(* CODESYS project SingleElevator.project

Project tree, tasks and I/O mapping:
  Device : CODESYS Control Win V3, 3S - Smart Software Solutions GmbH, version 3.5.18.0
    application Application
      libraries: Standard, 3.5.18.0 (System)
      task MainTask (cyclic, interval t#20ms, priority 1) calls GAs_Collector, Simulation, Policy
      task VISU_TASK (cyclic, interval 100 ms, priority 31) calls VisuElems.Visu_Prg
      global variables GVL
      visualisation Visualization
      program Simulation [ST]
      function block Cabin_GA [SFC]: Init_active, Ready_active, Busy_active, CabinUP_active, CabinUP_exit, CabinDown_exit, CabinDown_active, DoneHoming_active, DoneHoming_exit, HomingUp_active, HomingUp_exit, Step0_active, Step0_exit, ConteggioRampe_active, ConteggioDeck_active, Rallenta_active, Rallenta_exit, Fault_active, DoneCabin_active, FaultDeck_active, FaultDoneD_active, FaultDoneD_exit, FaultRamp_active, FaultDoneR_active, FaultDoneR_exit, FaultLimit_active, FaultLimit_exit, FaultDoneL_active, FaultDoneL_exit
      function block Doors_GA [SFC]: Init_active, Ready_active, Ready_exit, DoorOpening_active, DoorOpening_exit, SetDoneO_active, SetDoneO_exit, DoorClosing_active, DoorClosing_exit, SetDoneC_active, SetDoneC_exit
      function block HMI_GA [SFC]: Init_active, Ready_active, Ready_exit, LED_active, Chiamate_active, Destinazioni_active
      program Policy [SFC]: ChiusuraHoming_active, ChiusuraHoming_exit, Homing_active, Homing_exit, AperturaHoming_active, AperturaHoming_exit, Wait_Call_active, CalcoloDest_active, StopHMI_active, Chiudi_exit, Chiudi_active, Rallenta_active, AperturaEmergenza_active, Sali_active, Scendi_active, Sali_exit, Scendi_exit, Apri_exit, Apri_active
      program GAs_Collector [FBD]
  text list GlobalTextList
*)

// Device/Application/GVL

//{attribute 'qualified_only'}
VAR_GLOBAL
(* Elevator managing variables*)
	Open: BOOL;				(* Sensor: the door is fully open*)
	Closed: BOOL;			(* Sensor: the door is fully closed*)
	LimitDown: BOOL;		(* Sensor: lower limit sensor, if TRUE the lift has reached the lower limit*)
	LimitUp: BOOL;			(* Sensor: upper limit sensor, if TRUE the lift has reached the upper limit*)
	DeckSensor: BOOL;		(* Sensor: if TRUE the cab is in proximity of a deck*)
	RampSensor: BOOL;		(* Sensor: if TRUE the cab is in proximity of a ramp*)
	Presence :BOOL; 		(* Sensor: if TRUE something blocks the door photocell*)
	Emergency: BOOL;		(* Input: if TRUE the emergency button has been pressed*)

	Closing: BOOL;			(* Actuator: if TRUE the door starts closing*)
	Opening: BOOL;			(* Actuator: the door starts opening*)
	Motor_on: BOOL;			(* Actuator: if TRUE the lift pulley motor start moving*)
	Up: BOOL;				(* Actuator parameter: if TRUE the lift moves upward, downward otherwise*)
	Vel: BOOL;				(* Actuator parameter: motor speed, if TRUE high speed, low speed otherwise*)


	Current: INT;  			(* Visualization: variable used to storage the current deck*)
    Destination: INT;		(* Visualization: variable used to storage the the destination deck*)
	EmergencyVis: BOOL; 	(* Visualization: if TRUE the emergency light is turned on*)

	InitialDeck: INT := 1;	(* Only for simulation: variable used to define the initial deck*)
	InitCycle: BOOL := FALSE;(* Only for simulation: used to execute the instruction at the first cycle*)
	Height: INT;			(* Only for simulation: elevator height*)
	DeckRest: INT;        	(* Only for simulation: division rest for generating deck sensor*)
	Memory: INT;
	RampRest: INT;			(* Only for simulation: division rest for generating the ramp position*)
	MemoryR: INT;
	Door: INT;				(* Only for simulation: to visualize the closing of the door*)
	Displacement: INT;		(* Only for simulation: lift displacement, dependent on the motor speed*)

 (*Inputs: internal panel variables*)
	PG: BOOL;
	P1: BOOL;
	P2: BOOL;
	P3: BOOL;
	P4: BOOL;
	P5: BOOL;
	P6: BOOL;
	P7: BOOL;

(*Visualization: internal panel variables used to turn on the LED*)
	PGVis: BOOL;
	P1Vis: BOOL;
	P2Vis: BOOL;
	P3Vis: BOOL;
	P4Vis: BOOL;
	P5Vis: BOOL;
	P6Vis: BOOL;
	P7Vis: BOOL;

(*Inputs: external panel variables*)
	UpDeckG: BOOL;
	UpDeck1: BOOL;
	UpDeck2: BOOL;
	UpDeck3: BOOL;
	UpDeck4: BOOL;
	UpDeck5: BOOL;
	UpDeck6: BOOL;
	DownDeck7: BOOL;
	DownDeck6: BOOL;
	DownDeck5: BOOL;
	DownDeck4: BOOL;
	DownDeck3: BOOL;
	DownDeck2: BOOL;
	DownDeck1: BOOL;

(*Visualization: external panel variables used to turn on the LED*)
	UpDeckGVis: BOOL;
	UpDeck1Vis: BOOL;
	UpDeck2Vis: BOOL;
	UpDeck3Vis: BOOL;
	UpDeck4Vis: BOOL;
	UpDeck5Vis: BOOL;
	UpDeck6Vis: BOOL;
	DownDeck7Vis: BOOL;
	DownDeck6Vis: BOOL;
	DownDeck5Vis: BOOL;
	DownDeck4Vis: BOOL;
	DownDeck3Vis: BOOL;
	DownDeck2Vis: BOOL;
	DownDeck1Vis: BOOL;

(*Only for simulation: variables used to simulate the fault on deck sensor*)
	SensorG: BOOL;				(* if TRUE the magnetic information for deck G is lost and the deck sensor cannot become TRUE*)
	Sensor1: BOOL;				(* if TRUE the magnetic information for deck 1 is lost and the deck sensor cannot become TRUE*)
	Sensor2: BOOL;
	Sensor3: BOOL;
	Sensor4: BOOL;
	Sensor5: BOOL;
	Sensor6: BOOL;
	Sensor7: BOOL;
	FaultSensorAlarm: BOOL; 	(* Visulaization: if TRUE alerts the user of a deck sensor fault*)

(*Only for simulation: variables used to simulate the fault on ramp sensor*)
	RampGUp: BOOL;
	Ramp1Down: BOOL;
	Ramp1Up:BOOL;
	Ramp2Down: BOOL;
	Ramp2Up:BOOL;
	Ramp3Down: BOOL;
	Ramp3Up:BOOL;
	Ramp4Down: BOOL;
	Ramp4Up:BOOL;
	Ramp5Down: BOOL;
	Ramp5Up:BOOL;
	Ramp6Down: BOOL;
	Ramp6Up:BOOL;
	Ramp7Down: BOOL;
	FaultRampAlarm: BOOL; 		(* Visulaization: if TRUE alerts the user of a ramp sensor fault*)
	SensorGOK: BOOL;
	Sensor1OK: BOOL;
	Sensor2OK: BOOL;
	Sensor6OK: BOOL;
	Sensor3OK: BOOL;
	Sensor4OK: BOOL;
	Sensor5OK: BOOL;
	Sensor7OK: BOOL;
	RampGUpOK: BOOL;
	Ramp1DownOK: BOOL;
	Ramp1UpOK: BOOL;
	Ramp2DownOK: BOOL;
	Ramp2UpOK: BOOL;
	Ramp3DownOK: BOOL;
	Ramp3UpOK: BOOL;
	Ramp4DownOK: BOOL;
	Ramp4UpOK: BOOL;
	Ramp5DownOK: BOOL;
	Ramp5UpOK: BOOL;
	Ramp6DownOK: BOOL;
	Ramp6UpOK: BOOL;
	Ramp7DownOK: BOOL;
	Ramp7UpOK: BOOL;
	
	
	Cabin_GA_0: Cabin_GA;
	Doors_GA_0: Doors_GA;
	HMI_GA_0: HMI_GA;
END_VAR

// Device/Application/GAs_Collector
PROGRAM GAs_Collector
VAR
END_VAR

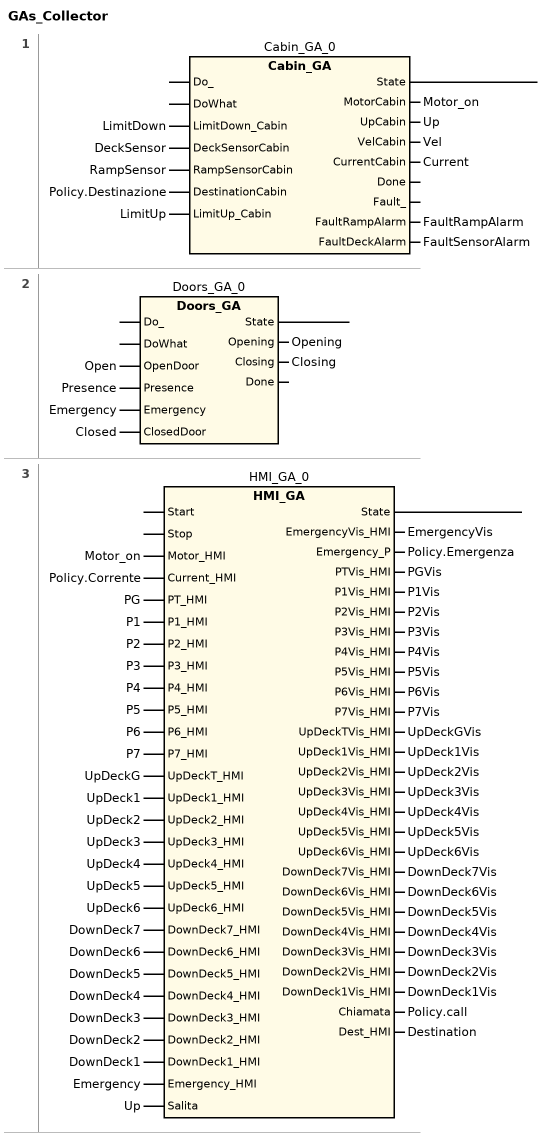
// NETWORK 1
Cabin_GA_0(
    LimitDown_Cabin := LimitDown,
    DeckSensorCabin := DeckSensor,
    RampSensorCabin := RampSensor,
    DestinationCabin := Policy.Destinazione,
    LimitUp_Cabin := LimitUp,
    MotorCabin => Motor_on,
    UpCabin => Up,
    VelCabin => Vel,
    CurrentCabin => Current,
    FaultRampAlarm => FaultRampAlarm,
    FaultDeckAlarm => FaultSensorAlarm); // Cabin_GA

// NETWORK 2
Doors_GA_0(
    OpenDoor := Open,
    Presence := Presence,
    Emergency := Emergency,
    ClosedDoor := Closed,
    Opening => Opening,
    Closing => Closing); // Doors_GA

// NETWORK 3
HMI_GA_0(
    Motor_HMI := Motor_on,
    Current_HMI := Policy.Corrente,
    PT_HMI := PG,
    P1_HMI := P1,
    P2_HMI := P2,
    P3_HMI := P3,
    P4_HMI := P4,
    P5_HMI := P5,
    P6_HMI := P6,
    P7_HMI := P7,
    UpDeckT_HMI := UpDeckG,
    UpDeck1_HMI := UpDeck1,
    UpDeck2_HMI := UpDeck2,
    UpDeck3_HMI := UpDeck3,
    UpDeck4_HMI := UpDeck4,
    UpDeck5_HMI := UpDeck5,
    UpDeck6_HMI := UpDeck6,
    DownDeck7_HMI := DownDeck7,
    DownDeck6_HMI := DownDeck6,
    DownDeck5_HMI := DownDeck5,
    DownDeck4_HMI := DownDeck4,
    DownDeck3_HMI := DownDeck3,
    DownDeck2_HMI := DownDeck2,
    DownDeck1_HMI := DownDeck1,
    Emergency_HMI := Emergency,
    Salita := Up,
    EmergencyVis_HMI => EmergencyVis,
    Emergency_P => Policy.Emergenza,
    PTVis_HMI => PGVis,
    P1Vis_HMI => P1Vis,
    P2Vis_HMI => P2Vis,
    P3Vis_HMI => P3Vis,
    P4Vis_HMI => P4Vis,
    P5Vis_HMI => P5Vis,
    P6Vis_HMI => P6Vis,
    P7Vis_HMI => P7Vis,
    UpDeckTVis_HMI => UpDeckGVis,
    UpDeck1Vis_HMI => UpDeck1Vis,
    UpDeck2Vis_HMI => UpDeck2Vis,
    UpDeck3Vis_HMI => UpDeck3Vis,
    UpDeck4Vis_HMI => UpDeck4Vis,
    UpDeck5Vis_HMI => UpDeck5Vis,
    UpDeck6Vis_HMI => UpDeck6Vis,
    DownDeck7Vis_HMI => DownDeck7Vis,
    DownDeck6Vis_HMI => DownDeck6Vis,
    DownDeck5Vis_HMI => DownDeck5Vis,
    DownDeck4Vis_HMI => DownDeck4Vis,
    DownDeck3Vis_HMI => DownDeck3Vis,
    DownDeck2Vis_HMI => DownDeck2Vis,
    DownDeck1Vis_HMI => DownDeck1Vis,
    Chiamata => Policy.call,
    Dest_HMI => Destination); // HMI_GA

END_PROGRAM

// Device/Application/Cabin_GA
FUNCTION_BLOCK Cabin_GA
VAR_INPUT
	Do_: BOOL;
	DoWhat: STRING;
	LimitDown_Cabin: BOOL;
	DeckSensorCabin: BOOL;
	RampSensorCabin: BOOL;
	DestinationCabin: INT;
	LimitUp_Cabin: BOOL;
END_VAR
VAR_OUTPUT
	State: STRING;
	MotorCabin: BOOL;
	UpCabin: BOOL;
	VelCabin: BOOL;
	CurrentCabin: INT;
	Done: BOOL;
	Fault_: BOOL;
	FaultRampAlarm: BOOL;
	FaultDeckAlarm: BOOL;
END_VAR
VAR
	N_rampe: INT;
	Dest: INT;
	Start: INT;
	i: INT; (*Rampe*)
	j: INT; (*Deck*)
	//k: INT; (*Rampe Aggiuntivo*)
	D_: BOOL;
	R_: BOOL;
	LUC: BOOL;
	LDC: BOOL;
END_VAR

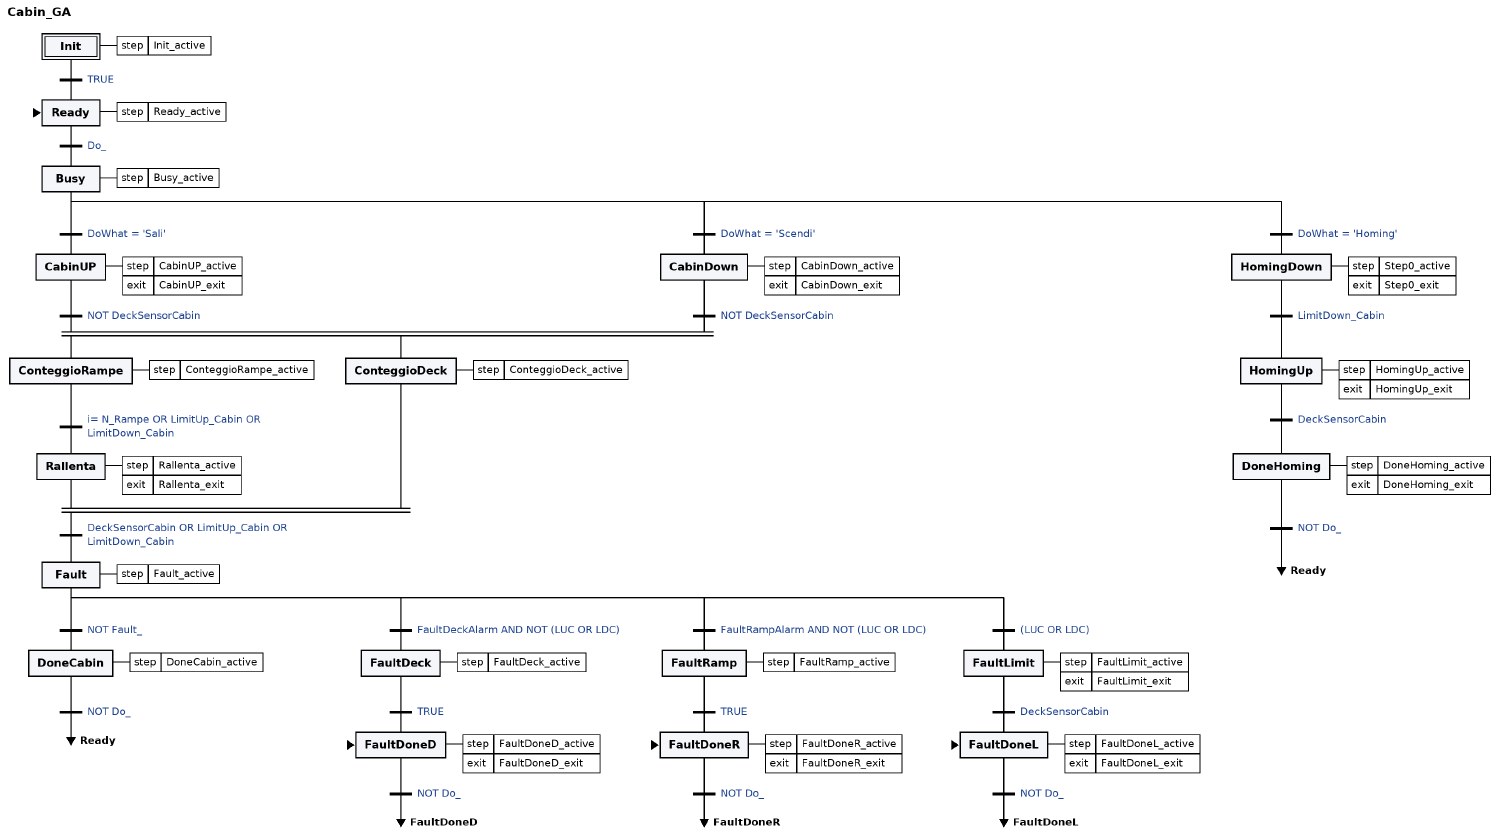
INITIAL_STEP Init:
    Init_active(N);  // step action
END_STEP
TRANSITION FROM Init TO Ready
    := TRUE;
END_TRANSITION
STEP Ready:
    Ready_active(N);  // step action
END_STEP
TRANSITION FROM Ready TO Busy
    := Do_;
END_TRANSITION
STEP Busy:
    Busy_active(N);  // step action
END_STEP
TRANSITION FROM Busy TO CabinUP
    := DoWhat = 'Sali';
END_TRANSITION
STEP CabinUP:
    CabinUP_active(N);  // step action
    CabinUP_exit(P0);  // exit action
END_STEP
TRANSITION FROM CabinUP TO (ConteggioRampe, ConteggioDeck)
    := NOT DeckSensorCabin;
END_TRANSITION
TRANSITION FROM Busy TO CabinDown
    := DoWhat = 'Scendi';
END_TRANSITION
STEP CabinDown:
    CabinDown_active(N);  // step action
    CabinDown_exit(P0);  // exit action
END_STEP
TRANSITION FROM CabinDown TO (ConteggioRampe, ConteggioDeck)
    := NOT DeckSensorCabin;
END_TRANSITION
TRANSITION FROM Busy TO HomingDown
    := DoWhat = 'Homing';
END_TRANSITION
STEP HomingDown:
    Step0_active(N);  // step action
    Step0_exit(P0);  // exit action
END_STEP
TRANSITION FROM HomingDown TO HomingUp
    := LimitDown_Cabin;
END_TRANSITION
STEP HomingUp:
    HomingUp_active(N);  // step action
    HomingUp_exit(P0);  // exit action
END_STEP
TRANSITION FROM HomingUp TO DoneHoming
    := DeckSensorCabin;
END_TRANSITION
STEP DoneHoming:
    DoneHoming_active(N);  // step action
    DoneHoming_exit(P0);  // exit action
END_STEP
TRANSITION FROM DoneHoming TO Ready
    := NOT Do_;
END_TRANSITION
STEP ConteggioRampe:
    ConteggioRampe_active(N);  // step action
END_STEP
TRANSITION FROM ConteggioRampe TO Rallenta
    := i= N_Rampe OR LimitUp_Cabin OR LimitDown_Cabin;
END_TRANSITION
STEP Rallenta:
    Rallenta_active(N);  // step action
    Rallenta_exit(P0);  // exit action
END_STEP
STEP ConteggioDeck:
    ConteggioDeck_active(N);  // step action
END_STEP
TRANSITION FROM (Rallenta, ConteggioDeck) TO Fault
    := DeckSensorCabin OR LimitUp_Cabin OR LimitDown_Cabin;
END_TRANSITION
STEP Fault:
    Fault_active(N);  // step action
END_STEP
TRANSITION FROM Fault TO DoneCabin
    := NOT Fault_;
END_TRANSITION
STEP DoneCabin:
    DoneCabin_active(N);  // step action
END_STEP
TRANSITION FROM DoneCabin TO Ready
    := NOT Do_;
END_TRANSITION
TRANSITION FROM Fault TO FaultDeck
    := FaultDeckAlarm AND NOT (LUC OR LDC);
END_TRANSITION
STEP FaultDeck:
    FaultDeck_active(N);  // step action
END_STEP
TRANSITION FROM FaultDeck TO FaultDoneD
    := TRUE;
END_TRANSITION
STEP FaultDoneD:
    FaultDoneD_active(N);  // step action
    FaultDoneD_exit(P0);  // exit action
END_STEP
TRANSITION FROM FaultDoneD TO FaultDoneD
    := NOT Do_;
END_TRANSITION
TRANSITION FROM Fault TO FaultRamp
    := FaultRampAlarm AND NOT (LUC OR LDC);
END_TRANSITION
STEP FaultRamp:
    FaultRamp_active(N);  // step action
END_STEP
TRANSITION FROM FaultRamp TO FaultDoneR
    := TRUE;
END_TRANSITION
STEP FaultDoneR:
    FaultDoneR_active(N);  // step action
    FaultDoneR_exit(P0);  // exit action
END_STEP
TRANSITION FROM FaultDoneR TO FaultDoneR
    := NOT Do_;
END_TRANSITION
TRANSITION FROM Fault TO FaultLimit
    := (LUC OR LDC);
END_TRANSITION
STEP FaultLimit:
    FaultLimit_active(N);  // step action
    FaultLimit_exit(P0);  // exit action
END_STEP
TRANSITION FROM FaultLimit TO FaultDoneL
    := DeckSensorCabin;
END_TRANSITION
STEP FaultDoneL:
    FaultDoneL_active(N);  // step action
    FaultDoneL_exit(P0);  // exit action
END_STEP
TRANSITION FROM FaultDoneL TO FaultDoneL
    := NOT Do_;
END_TRANSITION

ACTION Init_active:
State := 'Init';
END_ACTION

ACTION Ready_active:
State := 'Ready';
END_ACTION

ACTION Busy_active:
State := 'Busy';
END_ACTION

ACTION CabinUP_active:
MotorCabin := TRUE;
UpCabin := TRUE;
VelCabin :=FALSE;


N_rampe := (ABS(DestinationCabin - CurrentCabin)*2); (*Sensori di rampa attraversati*)
Dest := DestinationCabin;
Start:= CurrentCabin;
i:=0;
j:=0;
END_ACTION

ACTION CabinUP_exit:
VelCabin := TRUE;
END_ACTION

ACTION CabinDown_exit:
VelCabin := TRUE;
END_ACTION

ACTION CabinDown_active:
MotorCabin := TRUE;
UpCabin := FALSE;
VelCabin := FALSE;


N_rampe := (ABS(DestinationCabin - CurrentCabin)*2); (*Sensori di rampa attraversati*)
Dest := DestinationCabin;
Start:= CurrentCabin;
i:=0;
j:=0;
END_ACTION

ACTION DoneHoming_active:
Done :=TRUE;
END_ACTION

ACTION DoneHoming_exit:
Done := FALSE;
END_ACTION

ACTION HomingUp_active:
MotorCabin := TRUE;
UpCabin := TRUE;
VelCabin := FALSE;
END_ACTION

ACTION HomingUp_exit:
MotorCabin := FALSE;
CurrentCabin := 0;
END_ACTION

ACTION Step0_active:
MotorCabin := TRUE;
UpCabin := FALSE;
VelCabin := FALSE;
END_ACTION

ACTION Step0_exit:
MotorCabin := FALSE;
END_ACTION

ACTION ConteggioRampe_active:
IF RampSensorCabin = TRUE THEN
	IF R_ THEN
		i:=i+1;
		R_:=FALSE;
	END_IF
ELSE
	R_:=TRUE;
END_IF


IF Dest <> DestinationCabin THEN
	N_rampe := (ABS(DestinationCabin - Start)*2);
	Dest:=DestinationCabin;
END_IF
END_ACTION

ACTION ConteggioDeck_active:
IF DeckSensorCabin = TRUE THEN
	IF D_ THEN
		j:=j+1;
		D_:=FALSE;
		IF DoWhat = 'Sali' THEN
			CurrentCabin := CurrentCabin+1;
		ELSE
			CurrentCabin := CurrentCabin-1;
		END_IF
	END_IF
ELSE
	D_:=TRUE;
END_IF
END_ACTION

ACTION Rallenta_active:
VelCabin := FALSE;

IF RampSensor=TRUE THEN
	IF R_ THEN
		i:=i+1;
		R_:=FALSE;
	END_IF
ELSE
	R_:=TRUE;
END_IF
END_ACTION

ACTION Rallenta_exit:
MotorCabin := FALSE;
UpCabin := FALSE;
END_ACTION

ACTION Fault_active:
//Fault Deck/Fault Ramp
IF i<(2*j) AND NOT LUC AND NOT LDC THEN
	FaultRampAlarm :=TRUE;
	Fault_:=TRUE;
ELSIF i>(2*j) THEN
	FaultDeckAlarm :=TRUE;
	Fault_:=TRUE;
END_IF

//Fault Limit Up/Limit Down
IF LimitUp_Cabin THEN
	MotorCabin := TRUE;
	UpCabin:=FALSE;
	VelCabin := FALSE;
	LUC :=TRUE;
END_IF

IF LimitDown_Cabin THEN
	MotorCabin := TRUE;
	UpCabin:=TRUE;
	VelCabin := FALSE;
	LDC :=TRUE;
END_IF

IF LUC OR LDC THEN
	Fault_:=TRUE;
END_IF

//No Fault
IF i=2*j THEN
	Fault_:=FALSE;
END_IF
END_ACTION

ACTION DoneCabin_active:
Done := TRUE;
END_ACTION

ACTION FaultDeck_active:
IF DoWhat = 'Sali' THEN
	CurrentCabin := DestinationCabin+1;
ELSIF DoWhat = 'Scendi' THEN
	CurrentCabin := DestinationCabin-1;
END_IF

State := 'Fault_Deck';
DoWhat := 'Stop';
END_ACTION

ACTION FaultDoneD_active:
Done := TRUE;
END_ACTION

ACTION FaultDoneD_exit:
Done := FALSE;
END_ACTION

ACTION FaultRamp_active:
IF DoWhat = 'Sali' THEN
	CurrentCabin := DestinationCabin+1;
ELSIF DoWhat = 'Scendi' THEN
	CurrentCabin := DestinationCabin-1;
END_IF

State := 'Fault_Ramp';
DoWhat := 'Stop';
END_ACTION

ACTION FaultDoneR_active:
Done := TRUE;
END_ACTION

ACTION FaultDoneR_exit:
Done := FALSE;
END_ACTION

ACTION FaultLimit_active:
IF LUC THEN
	State := 'Fault_Deck';
END_IF

IF LDC THEN
	State:= 'Fault_Deck';
END_IF
END_ACTION

ACTION FaultLimit_exit:
MotorCabin := FALSE;
END_ACTION

ACTION FaultDoneL_active:
Done := TRUE;
END_ACTION

ACTION FaultDoneL_exit:
Done := false;
END_ACTION

END_FUNCTION_BLOCK

// Device/Application/Policy
PROGRAM Policy
VAR
	sync: BOOL;
	OpOk: BOOL;
	
	Destinazione: INT;
	Corrente: INT;
END_VAR

VAR_INPUT
	call: BOOL; 					//Presenza chiamate (origine: HMI)
	Emergenza: BOOL;				//Variabile di appoggio per Emergency (origine: HMI)
END_VAR

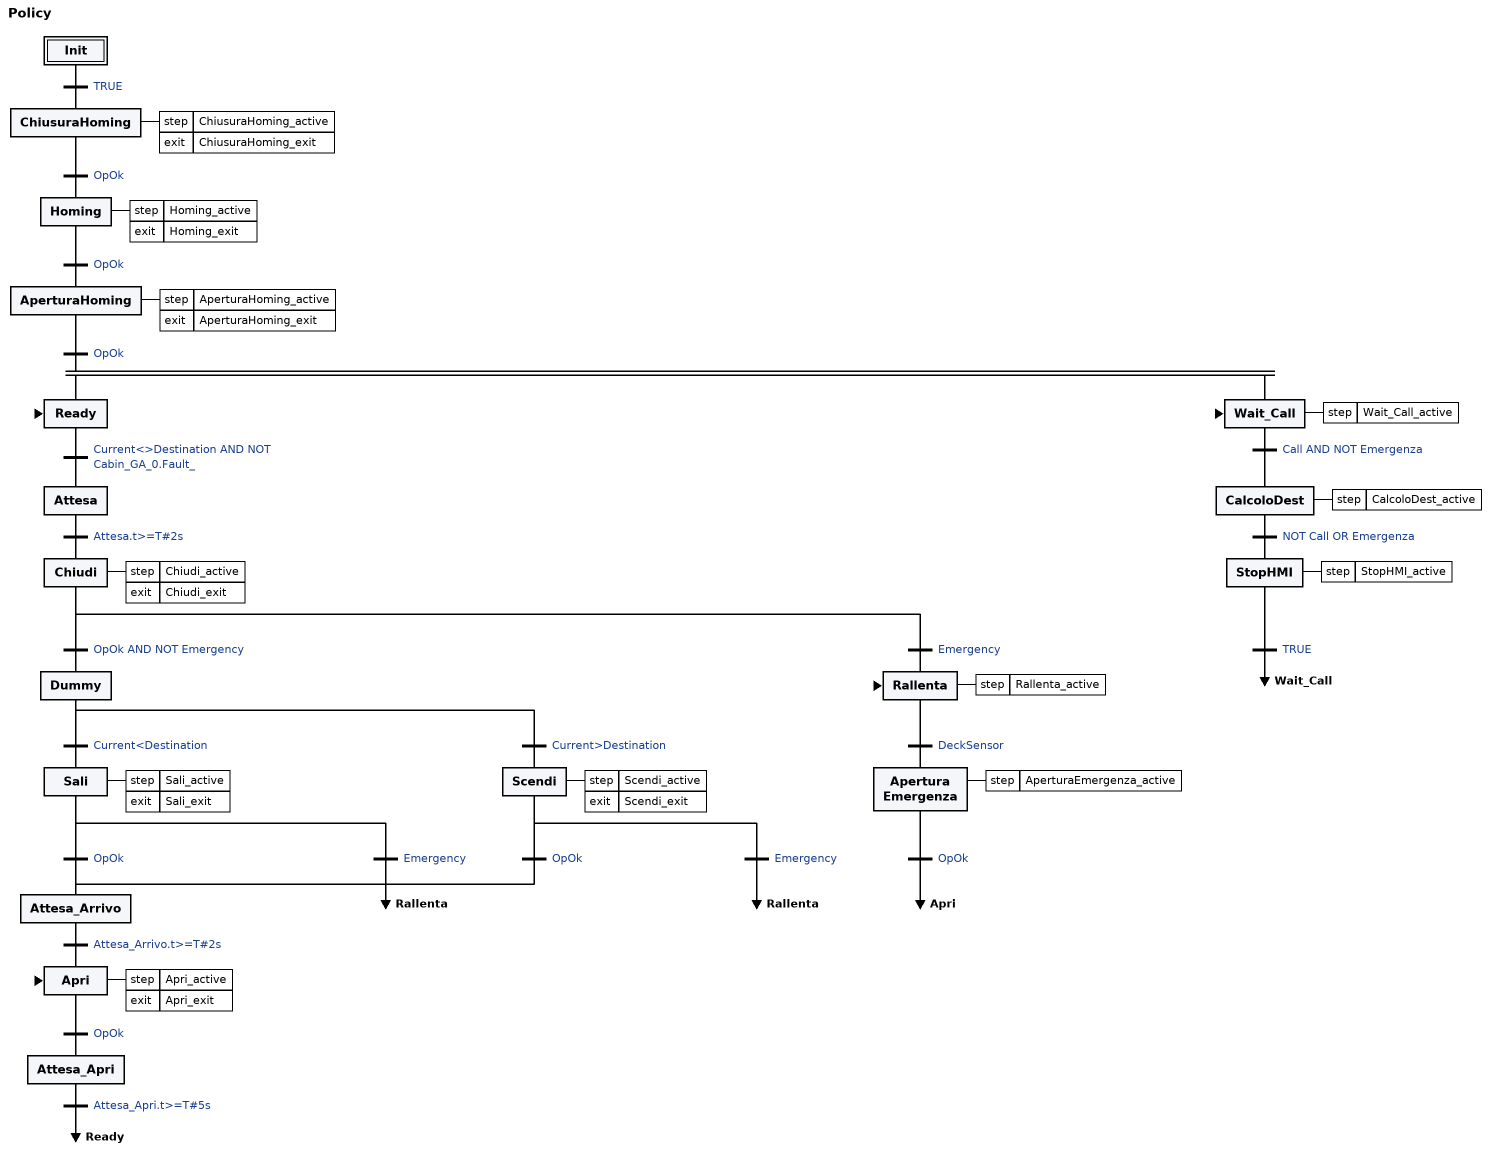
INITIAL_STEP Init:
END_STEP
TRANSITION FROM Init TO ChiusuraHoming
    := TRUE;
END_TRANSITION
STEP ChiusuraHoming:
    ChiusuraHoming_active(N);  // step action
    ChiusuraHoming_exit(P0);  // exit action
END_STEP
TRANSITION FROM ChiusuraHoming TO Homing
    := OpOk;
END_TRANSITION
STEP Homing:
    Homing_active(N);  // step action
    Homing_exit(P0);  // exit action
END_STEP
TRANSITION FROM Homing TO AperturaHoming
    := OpOk;
END_TRANSITION
STEP AperturaHoming:
    AperturaHoming_active(N);  // step action
    AperturaHoming_exit(P0);  // exit action
END_STEP
TRANSITION FROM AperturaHoming TO (Ready, Wait_Call)
    := OpOk;
END_TRANSITION
STEP Ready:
END_STEP
TRANSITION FROM Ready TO Attesa
    := Current<>Destination AND NOT Cabin_GA_0.Fault_;
END_TRANSITION
STEP Attesa:
END_STEP
TRANSITION FROM Attesa TO Chiudi
    := Attesa.t>=T#2s;
END_TRANSITION
STEP Chiudi:
    Chiudi_active(N);  // step action
    Chiudi_exit(P0);  // exit action
END_STEP
TRANSITION FROM Chiudi TO Dummy
    := OpOk AND NOT Emergency;
END_TRANSITION
STEP Dummy:
END_STEP
TRANSITION FROM Dummy TO Sali
    := Current<Destination;
END_TRANSITION
STEP Sali:
    Sali_active(N);  // step action
    Sali_exit(P0);  // exit action
END_STEP
TRANSITION FROM Sali TO Attesa_Arrivo
    := OpOk;
END_TRANSITION
TRANSITION FROM Sali TO Rallenta
    := Emergency;
END_TRANSITION
TRANSITION FROM Dummy TO Scendi
    := Current>Destination;
END_TRANSITION
STEP Scendi:
    Scendi_active(N);  // step action
    Scendi_exit(P0);  // exit action
END_STEP
TRANSITION FROM Scendi TO Attesa_Arrivo
    := OpOk;
END_TRANSITION
TRANSITION FROM Scendi TO Rallenta
    := Emergency;
END_TRANSITION
STEP Attesa_Arrivo:
END_STEP
TRANSITION FROM Attesa_Arrivo TO Apri
    := Attesa_Arrivo.t>=T#2s;
END_TRANSITION
STEP Apri:
    Apri_active(N);  // step action
    Apri_exit(P0);  // exit action
END_STEP
TRANSITION FROM Apri TO Attesa_Apri
    := OpOk;
END_TRANSITION
STEP Attesa_Apri:
END_STEP
TRANSITION FROM Attesa_Apri TO Ready
    := Attesa_Apri.t>=T#5s;
END_TRANSITION
TRANSITION FROM Chiudi TO Rallenta
    := Emergency;
END_TRANSITION
STEP Rallenta:
    Rallenta_active(N);  // step action
END_STEP
TRANSITION FROM Rallenta TO AperturaEmergenza
    := DeckSensor;
END_TRANSITION
STEP AperturaEmergenza:
    AperturaEmergenza_active(N);  // step action
END_STEP
TRANSITION FROM AperturaEmergenza TO Apri
    := OpOk;
END_TRANSITION
STEP Wait_Call:
    Wait_Call_active(N);  // step action
END_STEP
TRANSITION FROM Wait_Call TO CalcoloDest
    := Call AND NOT Emergenza;
END_TRANSITION
STEP CalcoloDest:
    CalcoloDest_active(N);  // step action
END_STEP
TRANSITION FROM CalcoloDest TO StopHMI
    := NOT Call OR Emergenza;
END_TRANSITION
STEP StopHMI:
    StopHMI_active(N);  // step action
END_STEP
TRANSITION FROM StopHMI TO Wait_Call
    := TRUE;
END_TRANSITION

ACTION ChiusuraHoming_active:
IF Presence = FALSE THEN
	IF Doors_GA_0.State = 'Ready' THEN
		Doors_GA_0.Do_:=TRUE;
		Doors_GA_0.DoWhat:='Chiudi';
	END_IF
END_IF

IF Doors_GA_0.Done AND Doors_GA_0.State='Busy' THEN
	Doors_GA_0.Do_:=FALSE;
	sync:=TRUE;
END_IF

OpOk:=sync AND Doors_GA_0.Done;
END_ACTION

ACTION ChiusuraHoming_exit:
sync:=FALSE;
OpOk:=FALSE;
END_ACTION

ACTION Homing_active:
IF Cabin_GA_0.State = 'Ready' THEN
	Cabin_GA_0.Do_:=TRUE;
	Cabin_GA_0.DoWhat:='Homing';
END_IF

IF Cabin_GA_0.Done AND Cabin_GA_0.State='Busy' THEN
	Cabin_GA_0.Do_:=FALSE;
	sync:=TRUE;
END_IF

OpOk:=sync AND Cabin_GA_0.Done;
END_ACTION

ACTION Homing_exit:
sync := FALSE;
OpOk := FALSE;
END_ACTION

ACTION AperturaHoming_active:
IF Doors_GA_0.State = 'Ready' THEN
	Doors_GA_0.Do_:=TRUE;
	Doors_GA_0.DoWhat:='Apri';
END_IF


IF Doors_GA_0.Done AND Doors_GA_0.State='Busy' THEN
	Doors_GA_0.Do_:=FALSE;
	sync:=TRUE;
END_IF

OpOk:=sync AND Doors_GA_0.Done;
END_ACTION

ACTION AperturaHoming_exit:
sync :=FALSE;
OpOk := FALSE;
END_ACTION

ACTION Wait_Call_active:
IF HMI_GA_0.State = 'Ready' THEN
	HMI_GA_0.Start:=TRUE;
	HMI_GA_0.Stop:=FALSE;
END_IF
END_ACTION

ACTION CalcoloDest_active:
Destinazione:=Destination;
Corrente:=Current;
END_ACTION

ACTION StopHMI_active:
IF HMI_GA_0.State = 'Busy' THEN
	HMI_GA_0.Start:=FALSE;
	HMI_GA_0.Stop:=TRUE;
END_IF
END_ACTION

ACTION Chiudi_exit:
sync := FALSE;
OpOk := FALSE;
END_ACTION

ACTION Chiudi_active:
IF Presence = FALSE THEN
	IF Doors_GA_0.State = 'Ready' THEN
		Doors_GA_0.Do_:=TRUE;
		Doors_GA_0.DoWhat:='Chiudi';
	END_IF
END_IF

IF Doors_GA_0.Done AND Doors_GA_0.State='Busy' THEN
	Doors_GA_0.Do_:=FALSE;
	sync:=TRUE;
END_IF

OpOk:=sync AND Doors_GA_0.Done;
END_ACTION

ACTION Rallenta_active:
Vel:= FALSE ;
END_ACTION

ACTION AperturaEmergenza_active:
Motor_on := FALSE;
IF Doors_GA_0.State = 'Ready' THEN
	Doors_GA_0.Do_:=TRUE;
	Doors_GA_0.DoWhat:='Apri';
END_IF


IF Doors_GA_0.Done AND Doors_GA_0.State='Busy' THEN
	Doors_GA_0.Do_:=FALSE;
	sync:=TRUE;
END_IF

OpOk:=sync AND Doors_GA_0.Done;
END_ACTION

ACTION Sali_active:
IF Cabin_GA_0.State='Ready' THEN
	Cabin_GA_0.Do_:=TRUE;
	Cabin_GA_0.DoWhat:='Sali';
END_IF

IF Cabin_GA_0.Done AND (Cabin_GA_0.State='Busy' OR Cabin_GA_0.State='Fault_Deck' OR Cabin_GA_0.State='Fault_Ramp') THEN
	Cabin_GA_0.Do_:=FALSE;
	sync:=TRUE;
END_IF

OpOk:=sync AND NOT Cabin_GA_0.Done;
END_ACTION

ACTION Scendi_active:
IF Cabin_GA_0.State='Ready' THEN
	Cabin_GA_0.Do_:=TRUE;
	Cabin_GA_0.DoWhat:='Scendi';
END_IF

IF Cabin_GA_0.Done AND (Cabin_GA_0.State='Busy' OR Cabin_GA_0.State='Fault_Deck' OR Cabin_GA_0.State='Fault_Ramp') THEN
	Cabin_GA_0.Do_:=FALSE;
	sync:=TRUE;
END_IF

OpOk:=sync AND NOT Cabin_GA_0.Done;
END_ACTION

ACTION Sali_exit:
sync:=FALSE;
OpOk:=FALSE;
END_ACTION

ACTION Scendi_exit:
sync:=FALSE;
OpOk:=FALSE;
END_ACTION

ACTION Apri_exit:
sync:=FALSE;
OpOk:=FALSE;
END_ACTION

ACTION Apri_active:
IF DeckSensor THEN	
	IF Doors_GA_0.State = 'Ready' THEN
		Doors_GA_0.Do_:=TRUE;
		Doors_GA_0.DoWhat:='Apri';
	END_IF


	IF Doors_GA_0.Done AND Doors_GA_0.State='Busy' THEN
		Doors_GA_0.Do_:=FALSE;
		sync:=TRUE;
	END_IF
END_IF

OpOk:=sync AND Doors_GA_0.Done;
END_ACTION

END_PROGRAM

// Device/Application/Doors_GA
FUNCTION_BLOCK Doors_GA
VAR_INPUT
	Do_: BOOL;
	DoWhat: STRING;
	OpenDoor: BOOL;
	Presence: BOOL;
	Emergency: BOOL;
	ClosedDoor: BOOL;
END_VAR
VAR_OUTPUT
	State: STRING;
	Opening: BOOL;
	Closing: BOOL;
	Done: BOOL;
END_VAR
VAR
END_VAR

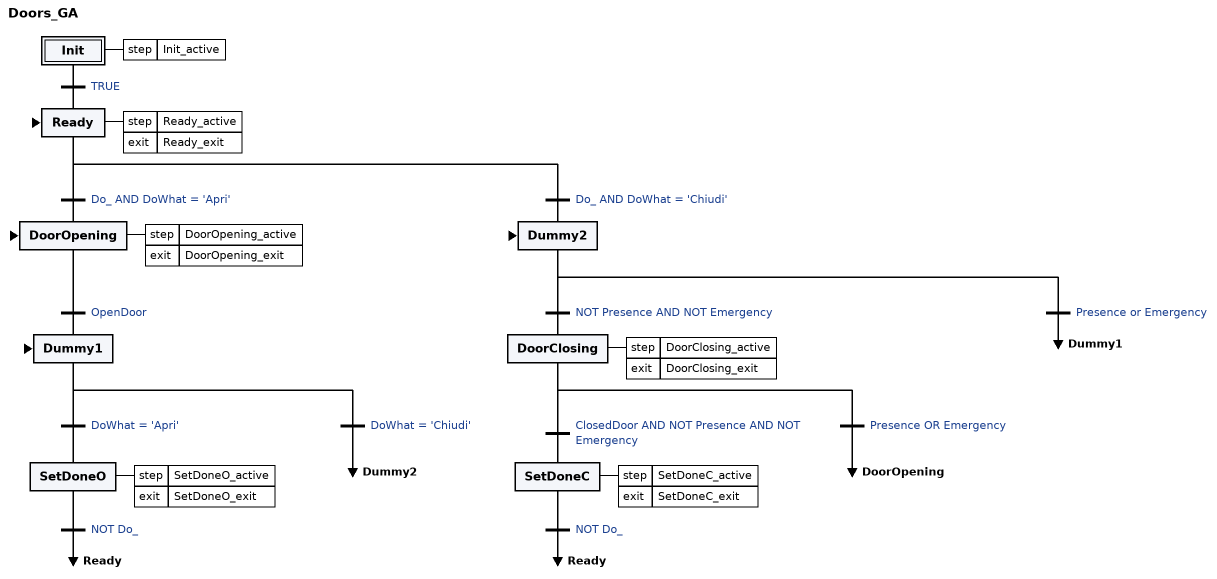
INITIAL_STEP Init:
    Init_active(N);  // step action
END_STEP
TRANSITION FROM Init TO Ready
    := TRUE;
END_TRANSITION
STEP Ready:
    Ready_active(N);  // step action
    Ready_exit(P0);  // exit action
END_STEP
TRANSITION FROM Ready TO DoorOpening
    := Do_ AND DoWhat = 'Apri';
END_TRANSITION
STEP DoorOpening:
    DoorOpening_active(N);  // step action
    DoorOpening_exit(P0);  // exit action
END_STEP
TRANSITION FROM DoorOpening TO Dummy1
    := OpenDoor;
END_TRANSITION
STEP Dummy1:
END_STEP
TRANSITION FROM Dummy1 TO SetDoneO
    := DoWhat = 'Apri';
END_TRANSITION
STEP SetDoneO:
    SetDoneO_active(N);  // step action
    SetDoneO_exit(P0);  // exit action
END_STEP
TRANSITION FROM SetDoneO TO Ready
    := NOT Do_;
END_TRANSITION
TRANSITION FROM Dummy1 TO Dummy2
    := DoWhat = 'Chiudi';
END_TRANSITION
TRANSITION FROM Ready TO Dummy2
    := Do_ AND DoWhat = 'Chiudi';
END_TRANSITION
STEP Dummy2:
END_STEP
TRANSITION FROM Dummy2 TO DoorClosing
    := NOT Presence AND NOT Emergency;
END_TRANSITION
STEP DoorClosing:
    DoorClosing_active(N);  // step action
    DoorClosing_exit(P0);  // exit action
END_STEP
TRANSITION FROM DoorClosing TO SetDoneC
    := ClosedDoor AND NOT Presence AND NOT Emergency;
END_TRANSITION
STEP SetDoneC:
    SetDoneC_active(N);  // step action
    SetDoneC_exit(P0);  // exit action
END_STEP
TRANSITION FROM SetDoneC TO Ready
    := NOT Do_;
END_TRANSITION
TRANSITION FROM DoorClosing TO DoorOpening
    := Presence OR Emergency;
END_TRANSITION
TRANSITION FROM Dummy2 TO Dummy1
    := Presence or Emergency;
END_TRANSITION

ACTION Init_active:
State := 'Init';
END_ACTION

ACTION Ready_active:
State := 'Ready';
END_ACTION

ACTION Ready_exit:
State := 'Busy';
END_ACTION

ACTION DoorOpening_active:
Opening := TRUE;
END_ACTION

ACTION DoorOpening_exit:
Opening := FALSE;
END_ACTION

ACTION SetDoneO_active:
Done := TRUE;
END_ACTION

ACTION SetDoneO_exit:
Done := FALSE;
END_ACTION

ACTION DoorClosing_active:
IF Presence = FALSE AND NOT ClosedDoor THEN 
	Closing := TRUE;
END_IF
END_ACTION

ACTION DoorClosing_exit:
Closing := FALSE;
END_ACTION

ACTION SetDoneC_active:
Done := TRUE;
END_ACTION

ACTION SetDoneC_exit:
Done := FALSE;
END_ACTION

END_FUNCTION_BLOCK

// Device/Application/HMI_GA
FUNCTION_BLOCK HMI_GA

VAR_OUTPUT
	State: STRING;
	EmergencyVis_HMI: BOOL;
	Emergency_P: BOOL;
	PTVis_HMI: BOOL;
	P1Vis_HMI: BOOL;
	P2Vis_HMI: BOOL;
	P3Vis_HMI: BOOL;
	P4Vis_HMI: BOOL;
	P5Vis_HMI: BOOL;
	P6Vis_HMI: BOOL;
	P7Vis_HMI: BOOL;
	UpDeckTVis_HMI: BOOL;
	UpDeck1Vis_HMI: BOOL;
	UpDeck2Vis_HMI: BOOL;
	UpDeck3Vis_HMI: BOOL;
	UpDeck4Vis_HMI: BOOL;
	UpDeck5Vis_HMI: BOOL;
	UpDeck6Vis_HMI: BOOL;
	DownDeck7Vis_HMI: BOOL;
	DownDeck6Vis_HMI: BOOL;
	DownDeck5Vis_HMI: BOOL;
	DownDeck4Vis_HMI: BOOL;
	DownDeck3Vis_HMI: BOOL;
	DownDeck2Vis_HMI: BOOL;
	DownDeck1Vis_HMI: BOOL;
	Chiamata: BOOL;
	Dest_HMI: INT;
END_VAR

VAR
	Interno: ARRAY[0..7] OF BOOL;
	Salire: ARRAY[0..7] OF BOOL;
	Scendere: ARRAY[0..7] OF BOOL;
	i: INT;
	
	Up_To: ARRAY [0..7] OF BOOL:= [FALSE, FALSE, FALSE, FALSE, FALSE, FALSE, FALSE, FALSE];
	Down_To: ARRAY [0..7] OF BOOL:= [FALSE, FALSE, FALSE, FALSE, FALSE, FALSE, FALSE, FALSE];
	
	flag: BOOL;
	w: INT;
	h: INT;
END_VAR

VAR_INPUT
	Start: BOOL;
	Stop: BOOL;
	Motor_HMI: BOOL;
	Current_HMI: INT;
	PT_HMI: BOOL;
	P1_HMI: BOOL;
	P2_HMI: BOOL;
	P3_HMI: BOOL;
	P4_HMI: BOOL;
	P5_HMI: BOOL;
	P6_HMI: BOOL;
	P7_HMI: BOOL;
	UpDeckT_HMI: BOOL;
	UpDeck1_HMI: BOOL;
	UpDeck2_HMI: BOOL;
	UpDeck3_HMI: BOOL;
	UpDeck4_HMI: BOOL;
	UpDeck5_HMI: BOOL;
	UpDeck6_HMI: BOOL;
	DownDeck7_HMI: BOOL;
	DownDeck6_HMI: BOOL;
	DownDeck5_HMI: BOOL;
	DownDeck4_HMI: BOOL;
	DownDeck3_HMI: BOOL;
	DownDeck2_HMI: BOOL;
	DownDeck1_HMI: BOOL;
	Emergency_HMI: BOOL;
	Salita: BOOL;
END_VAR

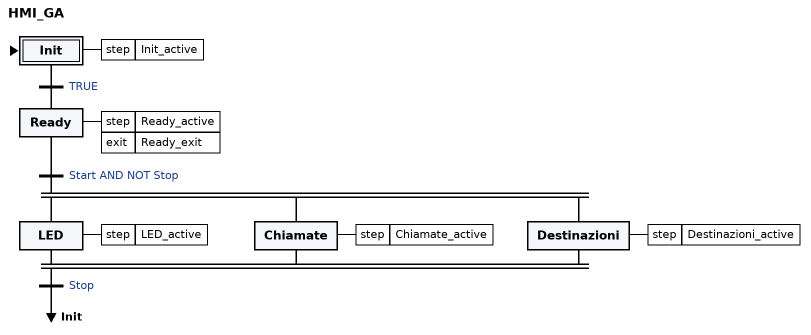
INITIAL_STEP Init:
    Init_active(N);  // step action
END_STEP
TRANSITION FROM Init TO Ready
    := TRUE;
END_TRANSITION
STEP Ready:
    Ready_active(N);  // step action
    Ready_exit(P0);  // exit action
END_STEP
TRANSITION FROM Ready TO (LED, Chiamate, Destinazioni)
    := Start AND NOT Stop;
END_TRANSITION
STEP LED:
    LED_active(N);  // step action
END_STEP
STEP Chiamate:
    Chiamate_active(N);  // step action
END_STEP
STEP Destinazioni:
    Destinazioni_active(N);  // step action
END_STEP
TRANSITION FROM (LED, Chiamate, Destinazioni) TO Init
    := Stop;
END_TRANSITION

ACTION Init_active:
State := 'Init';
END_ACTION

ACTION Ready_active:
State := 'Ready';
END_ACTION

ACTION Ready_exit:
State := 'Busy';
END_ACTION

ACTION LED_active:
//Accensione LED 
IF PT_HMI=TRUE THEN
	IF NOT(Motor_HMI=FALSE AND Current_HMI=0)THEN
		PTVis_HMI:=TRUE;
		Interno[0]:=TRUE;
	END_IF
ELSIF (Motor_HMI=FALSE AND Current_HMI=0) THEN
	PTVis_HMI:=FALSE;
	Interno[0]:=FALSE;
END_IF
	
IF P1_HMI=TRUE THEN
	IF NOT(Motor_HMI=FALSE AND Current_HMI=1) THEN
		P1Vis_HMI:=TRUE;
		Interno[1]:=TRUE;
	END_IF
ELSIF (Motor_HMI=FALSE AND Current_HMI=1) THEN
	P1Vis_HMI:=FALSE;
	Interno[1]:=FALSE;
END_IF
	
IF P2_HMI=TRUE THEN
	IF NOT(Motor_HMI=FALSE AND Current_HMI=2) THEN
		P2Vis_HMI:=TRUE;
		Interno[2]:=TRUE;
	END_IF
ELSIF (Motor_HMI=FALSE AND Current_HMI=2) THEN
	P2Vis_HMI:=FALSE;
	Interno[2]:=FALSE;
END_IF
	
IF P3_HMI=TRUE THEN
	IF NOT(Motor_HMI=FALSE AND Current_HMI=3) THEN
		P3Vis_HMI:=TRUE;
		Interno[3]:=TRUE;
	END_IF
ELSIF (Motor_HMI=FALSE AND Current_HMI=3) THEN
	P3Vis_HMI:=FALSE;
	Interno[3]:=FALSE;
END_IF

IF P4_HMI=TRUE THEN
	IF NOT(Motor_HMI=FALSE AND Current_HMI=4) THEN
		P4Vis_HMI:=TRUE;
		Interno[4]:=TRUE;
	END_IF
ELSIF (Motor_HMI=FALSE AND Current_HMI=4) THEN
	P4Vis_HMI:=FALSE;
	Interno[4]:=FALSE;
END_IF
	
IF P5_HMI=TRUE THEN
	IF NOT(Motor_HMI=FALSE AND Current_HMI=5) THEN
		P5Vis_HMI:=TRUE;
		Interno[5]:=TRUE;
	END_IF
ELSIF (Motor_HMI=FALSE AND Current_HMI=5) THEN
	P5Vis_HMI:=FALSE;
	Interno[5]:=FALSE;
END_IF
	
IF P6_HMI=TRUE THEN
	IF NOT(Motor_HMI=FALSE AND Current_HMI=6) THEN
		P6Vis_HMI:=TRUE;
		Interno[6]:=TRUE;
	END_IF
ELSIF (Motor_HMI=FALSE AND Current_HMI=6) THEN
	P6Vis_HMI:=FALSE;
	Interno[6]:=FALSE;
END_IF

IF P7_HMI=TRUE THEN
	IF NOT(Motor_HMI=FALSE AND Current_HMI=7) THEN
		P7Vis_HMI:=TRUE;
		Interno[7]:=TRUE;
	END_IF
ELSIF (Motor_HMI=FALSE AND Current_HMI=7) THEN
	P7Vis_HMI:=FALSE;
	Interno[7]:=FALSE;
END_IF
	
IF UpDeckT_HMI=TRUE THEN
	IF NOT(Motor_HMI=FALSE AND Current_HMI=0)THEN
		UpDeckTVis_HMI:=TRUE;
		Salire[0]:=TRUE;
	END_IF
ELSIF (Motor_HMI=FALSE AND Current_HMI=0) THEN
	UpDeckTVis_HMI:=FALSE;
	Salire[0]:=FALSE;
END_IF
	
IF UpDeck1_HMI=TRUE THEN
	IF NOT(Motor_HMI=FALSE AND Current_HMI=1) THEN
		UpDeck1Vis_HMI:=TRUE;
		Salire[1]:=TRUE;
	END_IF
ELSIF (Motor_HMI=FALSE AND Current_HMI=1) THEN
	UpDeck1Vis_HMI:=FALSE;
	Salire[1]:=FALSE;
END_IF

IF UpDeck2_HMI=TRUE THEN
	IF NOT(Motor_HMI=FALSE AND Current_HMI=2) THEN
		UpDeck2Vis_HMI:=TRUE;
		Salire[2]:=TRUE;
	END_IF
ELSIF (Motor_HMI=FALSE AND Current_HMI=2) THEN
	UpDeck2Vis_HMI:=FALSE;
	Salire[2]:=FALSE;
END_IF
	
IF UpDeck3_HMI=TRUE THEN
	IF NOT(Motor_HMI=FALSE AND Current_HMI=3) THEN
		UpDeck3Vis_HMI:=TRUE;
		Salire[3]:=TRUE;
	END_IF
ELSIF (Motor_HMI=FALSE AND Current_HMI=3) THEN
	UpDeck3Vis_HMI:=FALSE;
	Salire[3]:=FALSE;
END_IF
	
IF UpDeck4_HMI=TRUE THEN
	IF NOT(Motor_HMI=FALSE AND Current_HMI=4) THEN
		UpDeck4Vis_HMI:=TRUE;
		Salire[4]:=TRUE;
	END_IF
ELSIF (Motor_HMI=FALSE AND Current_HMI=4) THEN
	UpDeck4Vis_HMI:=FALSE;
	Salire[4]:=FALSE;
END_IF
	
IF UpDeck5_HMI=TRUE THEN
	IF NOT(Motor_HMI=FALSE AND Current_HMI=5) THEN
		UpDeck5Vis_HMI:=TRUE;
		Salire[5]:=TRUE;
	END_IF
ELSIF (Motor_HMI=FALSE AND Current_HMI=5) THEN
	UpDeck5Vis_HMI:=FALSE;
	Salire[5]:=FALSE;
END_IF
	
IF UpDeck6_HMI=TRUE THEN
	IF NOT(Motor_HMI=FALSE AND Current_HMI=6) THEN
		UpDeck6Vis_HMI:=TRUE;
		Salire[6]:=TRUE;
	END_IF
ELSIF (Motor_HMI=FALSE AND Current_HMI=6) THEN
	UpDeck6Vis_HMI:=FALSE;
	Salire[6]:=FALSE;
END_IF
	
IF DownDeck7_HMI=TRUE THEN
	IF NOT(Motor_HMI=FALSE AND Current_HMI=7)THEN
		DownDeck7Vis_HMI:=TRUE;
		Scendere[7]:=TRUE;
	END_IF
ELSIF (Motor_HMI=FALSE AND Current_HMI=7) THEN
	DownDeck7Vis_HMI:=FALSE;
	Scendere[7]:=FALSE;
END_IF
	
IF DownDeck6_HMI=TRUE THEN
	IF NOT(Motor_HMI=FALSE AND Current_HMI=6) THEN
		DownDeck6Vis_HMI:=TRUE;
		Scendere[6]:=TRUE;
	END_IF
ELSIF (Motor_HMI=FALSE AND Current_HMI=6) THEN
	DownDeck6Vis_HMI:=FALSE;
	Scendere[6]:=FALSE;
END_IF
	
IF DownDeck5_HMI=TRUE THEN
	IF NOT(Motor_HMI=FALSE AND Current_HMI=5) THEN
		DownDeck5Vis_HMI:=TRUE;
		Scendere[5]:=TRUE;
	END_IF
ELSIF (Motor_HMI=FALSE AND Current_HMI=5) THEN
	DownDeck5Vis_HMI:=FALSE;
	Scendere[5]:=FALSE;
END_IF
	
IF DownDeck4_HMI=TRUE THEN
	IF NOT(Motor_HMI=FALSE AND Current_HMI=4) THEN
		DownDeck4Vis_HMI:=TRUE;
		Scendere[4]:=TRUE;
	END_IF
ELSIF (Motor_HMI=FALSE AND Current_HMI=4) THEN
	DownDeck4Vis_HMI:=FALSE;
	Scendere[4]:=FALSE;
END_IF
	
IF DownDeck3_HMI=TRUE THEN
	IF NOT(Motor_HMI=FALSE AND Current_HMI=3) THEN
		DownDeck3Vis_HMI:=TRUE;
		Scendere[3]:=TRUE;
	END_IF
ELSIF (Motor_HMI=FALSE AND Current_HMI=3) THEN
	DownDeck3Vis_HMI:=FALSE;
	Scendere[3]:=FALSE;
END_IF
	
IF DownDeck2_HMI=TRUE THEN
	IF NOT(Motor_HMI=FALSE AND Current_HMI=2) THEN
		DownDeck2Vis_HMI:=TRUE;
		Scendere[2]:=TRUE;
	END_IF
ELSIF (Motor_HMI=FALSE AND Current_HMI=2) THEN
	DownDeck2Vis_HMI:=FALSE;
	Scendere[2]:=FALSE;
END_IF

IF DownDeck1_HMI=TRUE THEN
	IF NOT(Motor_HMI=FALSE AND Current_HMI=1)THEN
		DownDeck1Vis_HMI:=TRUE;
		Scendere[1]:=TRUE;
	END_IF
ELSIF (Motor_HMI=FALSE AND Current_HMI=1) THEN
	DownDeck1Vis_HMI:=FALSE;
	Scendere[1]:=FALSE;
END_IF
	
IF Emergency_HMI=TRUE THEN
	EmergencyVis_HMI:=TRUE;
	Emergency_P:=TRUE;
ELSE
	EmergencyVis_HMI:=FALSE;
	Emergency_P:=FALSE;
END_IF
END_ACTION

ACTION Chiamate_active:
//Lettura pulsanti
FOR i:=0 TO 7 BY 1 DO
	IF Interno[i] OR Salire[i] OR Scendere[i] THEN
		Chiamata:=TRUE;
	END_IF
END_FOR

//Riempimento Destinazioni In Salita e Destinazioni In Discesa
FOR i:=0 TO 7 BY 1 DO
	IF Interno[i] OR Salire[i] THEN
		Up_To[i]:=TRUE;
	ELSE
		Up_To[i]:=FALSE;
	END_IF
END_FOR

FOR i:=0 TO 7 BY 1 DO
	IF Interno[i] OR Scendere[i] THEN
		Down_To[i]:=TRUE;
	ELSE
		Down_To[i]:=FALSE;
	END_IF
END_FOR
END_ACTION

ACTION Destinazioni_active:
//Calcolo Destinazione
IF Salita OR flag THEN
	FOR w:=7 TO 0 BY (-1) DO
		IF Up_To[w] AND (w>Current_HMI OR NOT Motor_HMI) THEN		//Chiamate a Salire
			Dest_HMI:=w;
		END_IF
	END_FOR
	flag:=FALSE;
ELSIF NOT Motor_HMI OR NOT Salita OR NOT flag THEN
	FOR w:=0 TO 7 BY (1) DO
		IF Down_To[w] AND (w<Current_HMI OR NOT Motor_HMI) THEN		//Chiamate a Scendere
			Dest_HMI:=w;
			h:=0;
		ELSE
			h:=h+1;
			IF h=8 THEN														 
				flag:=TRUE;											 //Assenza di chiamate a Scendere
				h:=0;	
			END_IF
		END_IF
	END_FOR
END_IF

//Manovra di emergenza per fermata in sicurezza
IF Emergency_HMI THEN
    IF Dest_HMI<Current_HMI THEN
        Dest_HMI:=Current_HMI-1;
    ELSIF Dest_HMI>Current_HMI THEN
        Dest_HMI:=Current_HMI+1;
    END_IF
END_IF
END_ACTION

END_FUNCTION_BLOCK

// Device/Application/Simulation
PROGRAM Simulation
VAR
END_VAR

(* Initial position of the cab inside the hoistway. It is executed only at the first cycle.  *)
IF NOT GVL.InitCycle THEN
			GVL.InitCycle := TRUE ;
			GVL.Height := 20 * GVL.InitialDeck;
		    GVL.Door := 0;
			GVL.Current := GVL.Height / 20;
END_IF;

(* Elevator management, these instructions are executed each cycle time*)

(* Elevator door control. *)
IF GVL.Closing THEN
	GVL.Door := GVL.Door + 1;		(*Closing door management*)
	GVL.Open := FALSE;
END_IF

IF GVL.Door >= 60 THEN						(* Closed door limit*)
	GVL.Closed := TRUE;
END_IF

IF GVL.Opening THEN
	GVL.Door := GVL.Door - 1; 	(* Opening door management*)
	GVL.Closed := FALSE;
END_IF

IF GVL.Door <= 0 THEN							(* Open door limit*)
	GVL.Open := TRUE;
END_IF


(* Maximum and minimum management in the door simulation*)
IF GVL.Door < 0 THEN
	 GVL.Door := 0;
END_IF

IF GVL.Door > 60 THEN
	GVL.Door := 60;
END_IF


(* Control of the cab position inside the hostway. *)
(* Displacement definition for graphic visualization*)
IF GVL.Vel THEN 
	GVL.Displacement := 2;
ELSE 
	GVL.Displacement := 1;
END_IF


(* Height modification relying on direction and speed*)
IF GVL.Motor_on AND GVL.Up THEN
	GVL.Height := GVL.Height + GVL.Displacement;
	GVL.LimitDown := FALSE;
END_IF

IF GVL.Motor_on AND NOT GVL.Up THEN
	GVL.Height := GVL.Height - GVL.Displacement;
	GVL.LimitUp := FALSE;
END_IF


(* Limits for visualization*)
IF GVL.Height < -20 THEN
	GVL.Height := -20;
END_IF

IF GVL.Height > 160 THEN
	GVL.Height := 160;
END_IF

(* Limit sensors management*)
IF GVL.Height <= -10 THEN
	GVL.LimitDown := TRUE;
END_IF

IF GVL.Height >= 150 THEN
	 GVL.LimitUp := TRUE;
END_IF


(*-------------------------------------------------------------------*)
(*  Fault Management (Deck and Ramp Sensors)   *)
(*-------------------------------------------------------------------*)
(* Deck Sensor*)
(* Range of value where the deck sensor is active*)
IF ((GVL.Height >= -1) AND (GVL.Height <= 1)) THEN
	GVL.SensorGOK := TRUE;
ELSE  
	GVL.SensorGOK := FALSE;
END_IF

IF ((GVL.Height >= 20-1) AND (GVL.Height <= 20+1)) THEN
	GVL.Sensor1OK := TRUE;
ELSE  
	GVL.Sensor1OK := FALSE;
END_IF

IF ((GVL.Height >= 40-1) AND (GVL.Height <= 40+1)) THEN
	GVL.Sensor2OK := TRUE;
ELSE  
	GVL.Sensor2OK := FALSE;
END_IF

IF ((GVL.Height >= 60-1) AND (GVL.Height <= 60+1)) THEN
	GVL.Sensor3OK := TRUE;
ELSE  
	GVL.Sensor3OK := FALSE;
END_IF

IF ((GVL.Height >= 80-1) AND (GVL.Height <= 80+1)) THEN
	GVL.Sensor4OK := TRUE;
ELSE  
	GVL.Sensor4OK := FALSE;
END_IF

IF ((GVL.Height >= 100-1) AND (GVL.Height <= 100+1)) THEN
	GVL.Sensor5OK := TRUE;
ELSE   
	GVL.Sensor5OK := FALSE;
END_IF

IF ((GVL.Height >= 120-1) AND (GVL.Height <= 120+1)) THEN
	GVL.Sensor6OK := TRUE;
ELSE  
	GVL.Sensor6OK := FALSE;
END_IF

IF ((GVL.Height >= 140-1) AND (GVL.Height <= 140+1)) THEN
	GVL.Sensor7OK := TRUE;
ELSE  
	GVL.Sensor7OK := FALSE;
END_IF

GVL.DeckSensor := (GVL.SensorGOK AND NOT GVL.SensorG) OR
				    (GVL.Sensor1OK AND NOT GVL.Sensor1) OR
				    (GVL.Sensor2OK AND NOT GVL.Sensor2) OR
				    (GVL.Sensor3OK AND NOT GVL.Sensor3) OR
				    (GVL.Sensor4OK AND NOT GVL.Sensor4) OR
				    (GVL.Sensor5OK AND NOT GVL.Sensor5) OR
				    (GVL.Sensor6OK AND NOT GVL.Sensor6) OR
				    (GVL.Sensor7OK AND NOT GVL.Sensor7);

(* Ramp Sensor*)
(* Range of value where the ramp sensor is active*)
IF ((GVL.Height >= 5-1) AND (GVL.Height <= 5+1)) THEN
	GVL.RampGUpOK := TRUE;
ELSE 
	GVL.RampGUpOK := FALSE;
END_IF

(* Ramp close to deck 1*)
IF ((GVL.Height >= 15-1) AND (GVL.Height <= 15+1)) THEN
	GVL.Ramp1DownOK := TRUE;
ELSE 
	GVL.Ramp1DownOK := FALSE;
END_IF

IF ((GVL.Height >= 25-1) AND (GVL.Height <= 25+1)) THEN
	GVL.Ramp1UpOK := TRUE;
ELSE 
	GVL.Ramp1UpOK := FALSE;
END_IF

(* Ramp close to deck 2*)
IF ((GVL.Height >= 35-1) AND (GVL.Height <= 35+1)) THEN
	GVL.Ramp2DownOK := TRUE;
ELSE 
	GVL.Ramp2DownOK := FALSE;
END_IF

IF ((GVL.Height >= 45-1) AND (GVL.Height <= 45+1)) THEN
	GVL.Ramp2UpOK := TRUE;
ELSE 
	GVL.Ramp2UpOK := FALSE;
END_IF

(*Ramp close to deck  3*)
IF ((GVL.Height >= 55-1) AND (GVL.Height <= 55+1)) THEN
	GVL.Ramp3DownOK := TRUE;
ELSE 
	GVL.Ramp3DownOK := FALSE;
END_IF

IF ((GVL.Height >= 65-1) AND (GVL.Height <= 65+1)) THEN
	GVL.Ramp3UpOK := TRUE;
ELSE 
	GVL.Ramp3UpOK := FALSE;
END_IF

(* Ramp close to deck  4*)
IF ((GVL.Height >= 75-1) AND (GVL.Height <= 75+1)) THEN
	GVL.Ramp4DownOK := TRUE;
ELSE 
	GVL.Ramp4DownOK := FALSE;
END_IF

IF ((GVL.Height >= 85-1) AND (GVL.Height <= 85+1)) THEN
	GVL.Ramp4UpOK := TRUE;
ELSE 
	GVL.Ramp4UpOK:=FALSE;
END_IF

(* Ramp close to deck  5*)
IF ((GVL.Height >= 95-1) AND (GVL.Height <= 95+1)) THEN
	GVL.Ramp5DownOK := TRUE;
ELSE 
	GVL.Ramp5DownOK := FALSE;
END_IF

IF ((GVL.Height >= 105-1) AND (GVL.Height <= 105+1)) THEN
	GVL.Ramp5UpOK := TRUE;
ELSE
	GVL.Ramp5UpOK := FALSE;
END_IF

(* Ramp close to deck  6*)
IF ((GVL.Height >= 115-1) AND (GVL.Height <= 115+1)) THEN
	GVL.Ramp6DownOK := TRUE;
ELSE 
	GVL.Ramp6DownOK := FALSE;
END_IF

IF ((GVL.Height >= 125-1) AND (GVL.Height <= 125+1)) THEN
	GVL.Ramp6UpOK := TRUE;
ELSE 
	GVL.Ramp6UpOK := FALSE;
END_IF

(* Ramp close to deck  7*)
IF ((GVL.Height >= 135-1) AND (GVL.Height <= 135+1)) THEN
	GVL.Ramp7DownOK := TRUE;
ELSE 
	GVL.Ramp7DownOK := FALSE;
END_IF

GVL.RampSensor:=(GVL.RampGUpOK AND NOT GVL.RampGUp) OR 
								(GVL.Ramp1DownOK AND NOT GVL.Ramp1Down ) OR 
								(GVL.Ramp1UpOK AND NOT GVL.Ramp1Up ) OR
								(GVL.Ramp2DownOK AND NOT GVL.Ramp2Down ) OR 
								(GVL.Ramp2UpOK AND NOT GVL.Ramp2Up ) OR
								(GVL.Ramp3DownOK AND NOT GVL.Ramp3Down ) OR
 								(GVL.Ramp3UpOK AND NOT GVL.Ramp3Up ) OR
								(GVL.Ramp4DownOK AND NOT GVL.Ramp4Down ) OR
 								(GVL.Ramp4UpOK AND NOT GVL.Ramp4Up ) OR
								(GVL.Ramp5DownOK AND NOT GVL.Ramp5Down ) OR
 								(GVL.Ramp5UpOK AND NOT GVL.Ramp5Up ) OR
								(GVL.Ramp6DownOK AND NOT GVL.Ramp6Down ) OR
								(GVL.Ramp6UpOK AND NOT GVL.Ramp6Up ) OR
								(GVL.Ramp7DownOK AND NOT GVL.Ramp7Down );

END_PROGRAM

// Device/Application/Visualization
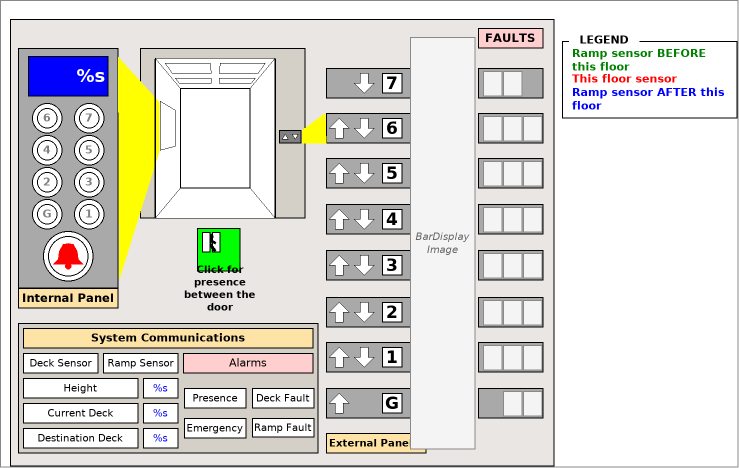
VISUALIZATION Visualization  // 739x468
    Rectangle (10,19 544x447)
    Rectangle (197,228 43x43), colour toggle: GVL.Presence
    Rectangle (18,323 300x130)
    Rectangle (326,433 100x20), "External Panels"
    Rectangle (326,342 100x30)
    Rectangle (382,347 20x20), "1"
    Polygon (354,357) (360,357) (360,347) (368,347) (368,357) (374,357) (364,367), colour toggle: GVL.DownDeck1Vis
        tap GVL.DownDeck1
    Polygon (329,357) (335,357) (335,367) (343,367) (343,357) (349,357) (339,347), colour toggle: GVL.UpDeck1Vis
        tap GVL.UpDeck1
    Rectangle (326,297 100x30)
    Rectangle (382,302 20x20), "2"
    Polygon (354,312) (360,312) (360,302) (368,302) (368,312) (374,312) (364,322), colour toggle: GVL.DownDeck2Vis
        tap GVL.DownDeck2
    Polygon (329,312) (335,312) (335,322) (343,322) (343,312) (349,312) (339,302), colour toggle: GVL.UpDeck2Vis
        tap GVL.UpDeck2
    Rectangle (326,250 100x30)
    Rectangle (382,255 20x20), "3"
    Polygon (354,265) (360,265) (360,255) (368,255) (368,265) (374,265) (364,275), colour toggle: GVL.DownDeck3Vis
        tap GVL.DownDeck3
    Polygon (329,265) (335,265) (335,275) (343,275) (343,265) (349,265) (339,255), colour toggle: GVL.UpDeck3Vis
        tap GVL.UpDeck3
    Rectangle (326,204 100x30)
    Rectangle (382,209 20x20), "4"
    Polygon (354,219) (360,219) (360,209) (368,209) (368,219) (374,219) (364,229), colour toggle: GVL.DownDeck4Vis
        tap GVL.DownDeck4
    Polygon (329,219) (335,219) (335,229) (343,229) (343,219) (349,219) (339,209), colour toggle: GVL.UpDeck4Vis
        tap GVL.UpDeck4
    Rectangle (326,158 100x30)
    Rectangle (382,163 20x20), "5"
    Polygon (354,173) (360,173) (360,163) (368,163) (368,173) (374,173) (364,183), colour toggle: GVL.DownDeck5Vis
        tap GVL.DownDeck5
    Polygon (329,173) (335,173) (335,183) (343,183) (343,173) (349,173) (339,163), colour toggle: GVL.UpDeck5Vis
        tap GVL.UpDeck5
    Rectangle (326,113 100x30)
    Rectangle (382,118 20x20), "6"
    Polygon (354,128) (360,128) (360,118) (368,118) (368,128) (374,128) (364,138), colour toggle: GVL.DownDeck6Vis
        tap GVL.DownDeck6
    Polygon (329,128) (335,128) (335,138) (343,138) (343,128) (349,128) (339,118), colour toggle: GVL.UpDeck6Vis
        tap GVL.UpDeck6
    Rectangle (326,68 100x30)
    Rectangle (382,73 20x20), "7"
    Polygon (354,83) (360,83) (360,73) (368,73) (368,83) (374,83) (364,93), colour toggle: GVL.DownDeck7Vis
        tap GVL.DownDeck7
    Rectangle (326,388 100x30)
    Rectangle (382,393 20x20), "G"
    Polygon (329,403) (335,403) (335,413) (343,413) (343,403) (349,403) (339,393), colour toggle: GVL.UpDeckGVis
        tap GVL.UpDeckG
    RoundedRectangle (18,48 100x240)
    Rectangle (18,288 100x20), "Internal Panel"
    Ellipse (74,199 30x30), colour toggle: GVL.P1Vis
    Ellipse (79,204 20x20), "1"
        tap GVL.P1
    Ellipse (32,199 30x30), colour toggle: GVL.PGVis
    Ellipse (37,204 20x20), "G"
        tap GVL.PG
    Ellipse (74,167 30x30), colour toggle: GVL.P3Vis
    Ellipse (79,172 20x20), "3"
        tap GVL.P3
    Ellipse (32,167 30x30), colour toggle: GVL.P2Vis
    Ellipse (37,172 20x20), "2"
        tap GVL.P2
    Ellipse (74,135 30x30), colour toggle: GVL.P5Vis
    Ellipse (79,140 20x20), "5"
        tap GVL.P5
    Ellipse (32,135 30x30), colour toggle: GVL.P4Vis
    Ellipse (37,140 20x20), "4"
        tap GVL.P4
    Ellipse (74,103 30x30), colour toggle: GVL.P7Vis
    Ellipse (79,108 20x20), "7"
        tap GVL.P7
    Ellipse (32,103 30x30), colour toggle: GVL.P6Vis
    Ellipse (37,108 20x20), "6"
        tap GVL.P6
    Rectangle (28,56 80x40), "%s", text variable: GVL.Destination
    Ellipse (43,231 50x50), tooltip "EMERGENCY", colour toggle: GVL.Emergency
    Group (48,236 40x40)
        toggle GVL.Emergency
        Ellipse (0,0 40x40), tooltip "EMERGENCY"
        Polygon (5,28) (10,23) (11,15) (15,8) (20,7) (25,8) (29,15) (30,23) (35,28)
        Ellipse (17,27 6x6)
    Polygon (35,72) (45,62) (55,72), colour toggle: GVL.Motor_on AND GVL.Up
    Polygon (35,80) (45,90) (55,80), colour toggle: GVL.Motor_on AND NOT GVL.Up
    Group (140,48 165x170)
        Rectangle (0,0 165x170)
        Rectangle (15,10 120x160)
        Polygon (40,40) (15,10) (135,10) (110,40)
        Rectangle (40,40 70x100)
        Polygon (15,170) (40,140) (110,140) (135,170)
        Polygon (20,102) (20,53) (35,62) (35,98)
        Polygon (79,35) (79,30) (115,30) (111,35)
        Polygon (39,35) (35,30) (71,30) (71,35)
        Polygon (32,25) (25,15) (70,15) (71,25)
        Polygon (79,25) (80,15) (125,15) (118,25)
        Group (139,82 22x13)
            Rectangle (0,0 22x13)
            Polygon (3,9) (6,4) (9,9)
            Polygon (13,4) (16,9) (19,4)
    BarDisplayImage (410,37 65x412), value: GVL.Height, style: BarDisplayImage-Gray, scale format: %.0f, scale -20..160
        p3451962224: VisuNativeControl.IP_Offline.Browser
    Rectangle (478,68 65x30)
    Rectangle (478,342 65x30)
    Rectangle (478,297 65x30)
    Rectangle (478,250 65x30)
    Rectangle (478,204 65x30)
    Rectangle (478,158 65x30)
    Rectangle (478,113 65x30)
    Rectangle (478,388 65x30)
    RockerSwitch (483,345 19x25), variable: GVL.Ramp1Down, behaviour: TOGGLE, style: Switch-RockerSwitch-Green
    RockerSwitch (503,345 19x25), variable: GVL.Sensor1, behaviour: TOGGLE, style: Switch-RockerSwitch-Red
    RockerSwitch (523,345 19x25), variable: GVL.Ramp1Up, behaviour: TOGGLE, style: Switch-RockerSwitch-Blue
    RockerSwitch (483,300 19x25), variable: GVL.Ramp2Down, behaviour: TOGGLE, style: Switch-RockerSwitch-Green
    RockerSwitch (503,300 19x25), variable: GVL.Sensor2, behaviour: TOGGLE, style: Switch-RockerSwitch-Red
    RockerSwitch (523,300 19x25), variable: GVL.Ramp2Up, behaviour: TOGGLE, style: Switch-RockerSwitch-Blue
    RockerSwitch (483,253 19x25), variable: GVL.Ramp3Down, behaviour: TOGGLE, style: Switch-RockerSwitch-Green
    RockerSwitch (503,253 19x25), variable: GVL.Sensor3, behaviour: TOGGLE, style: Switch-RockerSwitch-Red
    RockerSwitch (523,253 19x25), variable: GVL.Ramp3Up, behaviour: TOGGLE, style: Switch-RockerSwitch-Blue
    RockerSwitch (483,207 19x25), variable: GVL.Ramp4Down, behaviour: TOGGLE, style: Switch-RockerSwitch-Green
    RockerSwitch (503,207 19x25), variable: GVL.Sensor4, behaviour: TOGGLE, style: Switch-RockerSwitch-Red
    RockerSwitch (523,207 19x25), variable: GVL.Ramp4Up, behaviour: TOGGLE, style: Switch-RockerSwitch-Blue
    RockerSwitch (483,161 19x25), variable: GVL.Ramp5Down, behaviour: TOGGLE, style: Switch-RockerSwitch-Green
    RockerSwitch (503,161 19x25), variable: GVL.Sensor5, behaviour: TOGGLE, style: Switch-RockerSwitch-Red
    RockerSwitch (523,161 19x25), variable: GVL.Ramp5Up, behaviour: TOGGLE, style: Switch-RockerSwitch-Blue
    RockerSwitch (483,116 19x25), variable: GVL.Ramp6Down, behaviour: TOGGLE, style: Switch-RockerSwitch-Green
    RockerSwitch (503,116 19x25), variable: GVL.Sensor6, behaviour: TOGGLE, style: Switch-RockerSwitch-Red
    RockerSwitch (523,116 19x25), variable: GVL.Ramp6Up, behaviour: TOGGLE, style: Switch-RockerSwitch-Blue
    RockerSwitch (483,71 19x25), variable: GVL.Ramp7Down, behaviour: TOGGLE, style: Switch-RockerSwitch-Green
    RockerSwitch (503,71 19x25), variable: GVL.Sensor7, behaviour: TOGGLE, style: Switch-RockerSwitch-Red
    RockerSwitch (503,391 19x25), variable: GVL.SensorG, behaviour: TOGGLE, style: Switch-RockerSwitch-Red
    RockerSwitch (523,391 19x25), variable: GVL.RampGUp, behaviour: TOGGLE, style: Switch-RockerSwitch-Blue
    Rectangle (478,28 65x20), "FAULTS"
    Polygon (302,130) (325,113) (326,143) (302,143), invisible if: (GVL.Closing OR GVL.Opening) OR GVL.Closed
    Polygon (118,57) (159,102) (159,151) (119,279), invisible if: (GVL.Closing OR GVL.Opening) OR GVL.Closed
    Rectangle (155,58 0x160)
        p3528305787: GVL.Door
    Rectangle (275,58 0x160)
        p3528305787: -GVL.Door
    Rectangle (23,328 290x20), "System Communications"
    Rectangle (183,353 130x20), "Alarms"
    Rectangle (23,353 75x20), "Deck Sensor", colour toggle: GVL.DeckSensor
    Rectangle (143,378 35x20), "%s", text variable: GVL.Height
    Rectangle (184,388 62x20), "Presence", colour toggle: GVL.Presence
    Rectangle (103,353 75x20), "Ramp Sensor", colour toggle: GVL.RampSensor
    Rectangle (143,403 35x20), "%s", text variable: GVL.Current
    Rectangle (143,428 35x20), "%s", text variable: GVL.Destination
    Rectangle (252,388 62x20), "Deck Fault", colour toggle: GVL.FaultSensorAlarm
    Rectangle (184,418 62x20), "Emergency", colour toggle: GVL.EmergencyVis
    Rectangle (252,418 62x19), "Ramp Fault", colour toggle: GVL.FaultRampAlarm
    Rectangle (23,378 115x20), "Height"
    Rectangle (23,403 115x20), "Current Deck"
    Rectangle (23,428 115x20), "Destination Deck"
    Group (562,25 175x93)
        Rectangle (0,16 175x77)
        Rectangle (7,39 160x30), "This floor sensor"
        Rectangle (7,59 160x30), "Ramp sensor AFTER this floor"
        Rectangle (7,0 70x30), "LEGEND"
        Rectangle (7,20 160x30), "Ramp sensor BEFORE this floor"
    Group (202,232 33x34)
        toggle GVL.Presence
        Rectangle (10,0 8x20)
        Polygon (5,10) (12,20) (14,18) (5,6)
        Ellipse (6,2 5x5)
        Polygon (4,8) (13,12) (14,10) (4,4)
        Rectangle (0,0 8x20)
    Rectangle (169,273 102x31), "Click for presence between the door"
END_VISUALIZATION
